(* IEC 61131-3 sources: SRCI_CLIENT_PLC/RobotLibrary/Library/Constants, 2 files *)

(* ---- RobotLibraryConstants.st ---- *)
{attribute 'qualified_only'}
// -------------------------------------------------------------------------
//  SRCI Robot Library
// -------------------------------------------------------------------------
//
//  Object:      RobotLibraryConstants
//  Author:      Thorsten Brach
//  Date:        2024-06-01
//
//  Description:
//
//
//  Copyright:
//    (C) 2024 Thorsten Brach. All rights reserved
//             Licensed under the MIT License.
//
//  Disclaimer:
//    This project is provided without any guarantee and can be used for
//    private and commercial purposes. Any use is at the user’s
//    own risk and responsibility.
//
// -------------------------------------------------------------------------
VAR_GLOBAL CONSTANT
  /// Version of SRCI specification
  /// Bit 0-4 : Minor version = Features        (0..31)
  /// Bit 5-7 : Major version = Breaking change (0..07)
  SRCIVersion             : VersionStruct := ( MajorVersion := 1, MinorVersion := 5, PatchVersion := 0); // ST-FIX PLC library still says 1.3.0, but implements SRCI 1.5 (SDK: SRCI_VERSION 1.5)
  /// Version of the PLC library
  PLCLibraryVersion       : VersionStruct := ( MajorVersion := 1, MinorVersion := 5, PatchVersion := 7); // ST-FIX F166: the constant was not counted up (1.5.4 in library 1.5.5.0); now the release 1.5.7
  /// Minimal axes group ID
  AXES_GROUP_ID_MIN       : BYTE := 0;
  /// Maximal axes groups ID
  AXES_GROUP_ID_MAX       : BYTE := 15;
  /// OK = 0
  OK                      : DINT := 0;
  /// Running = 1
  RUNNING                 : DINT := 1;
  /// HasError = -1
  HAS_ERROR               : DINT := -1;
  /// Null pointer
  XNULL                   : DWORD := 0;
  /// Null pointer
  NULL_POINTER            : POINTER TO BYTE := 0;
  /// Real conversion factor ( REAL * 100 -> TO_INT )
  REAL_CONVERSION_FACTOR  : REAL := 100;
  /// Active command
  ACTIVE_CMD              : UDINT := 1;
  /// Buffered command
  BUFFER_CMD              : UDINT := 2;
  /// Maximal length of additional text
  MAX_ADD_TEXT_LENGTH     : DINT := 40;
  /// ST-FIX F108: characters of a log line per ReadServerLog response (SRCI SDK 1.1: 179;
  /// spec table 6-124: 187)
  SERVER_LOG_CONTENT_MAX  : DINT := 179;
  /// Upper index of the cyclic sub program data: 26 bytes (spec table 5-88, 6-711)
  /// ST-FIX F179: one constant for all arrays of the cyclic sub program data
  CYCLIC_SUB_PROGRAM_DATA_MAX : DINT := 25;
 END_VAR

(* ---- RobotLibraryDefines.st ---- *)
{attribute 'qualified_only'}
// -------------------------------------------------------------------------
//  SRCI Robot Library
// -------------------------------------------------------------------------
//
//  Object:      RobotLibraryDefines
//  Author:      Thorsten Brach
//  Date:        2024-06-01
//
//  Description:
//
//
//  Copyright:
//    (C) 2024 Thorsten Brach. All rights reserved
//             Licensed under the MIT License.
//
//  Disclaimer:
//    This project is provided without any guarantee and can be used for
//    private and commercial purposes. Any use is at the user’s
//    own risk and responsibility.
//
// -------------------------------------------------------------------------
VAR_GLOBAL
  /// Maximal length of type name
  MaxTypeNameLength  : INT;
END_VAR
